Staubli VAL3: aioItem.dtx

public string sComment
public aio aAio
